--- program FrameL (robot ABB IRB 1300-10/1.15) ---
  Smooth(1)
  Set speed (1000.0 mm/s)
  Set Ref.: FrameL
  Set Tool: Generic Paint Sprayer
  Show Generic Paint Sprayer
  MoveJ 1 to (-13.41, 234.2, 55.45) mm, rotated rx -20.36 ry -7.23 rz -177.33 deg; joints [77.348, 64.389, -177.634, -26.013, 92.152, 94.605, 581.087, 3508.568, 217.224]
  MoveL 2 to (-13.41, 234.2, 55.45) mm, rotated rx -20.36 ry -7.23 rz -177.33 deg; joints [77.348, 64.389, -177.634, -26.013, 92.152, 94.605, 581.087, 3508.568, 217.224]
  MoveL 3 to (0, 200, 148.46) mm, rotated rx -20.36 ry -7.23 rz -177.33 deg; joints [77.348, 64.389, -177.634, -26.013, 92.152, 94.605, 594.495, 3417.935, 257.297]
  MoveL 4 to (0, 200, 148.46) mm, rotated rx -20.36 ry -7.23 rz -177.33 deg; joints [77.348, 64.389, -177.634, -26.013, 92.152, 94.605, 594.495, 3417.935, 257.297]
  Set speed (20.0 mm/s)
  MoveL 5 to (0, 100, 118.49) mm, rotated rx -13.25 ry -10.31 rz -177.59 deg; joints [77.348, 64.389, -177.469, -28.671, 97.668, 89.928, 571.606, 3460.539, 412.588]
  MoveL 6 to (0, 0, 100.67) mm, rotated rx -6.84 ry -13.03 rz -178.45 deg; joints [77.348, 64.389, -174.962, -31.186, 100.159, 86.521, 548.69, 3498.334, 553.088]
  Set speed (1000.0 mm/s)
  MoveL 7 to (0, 0, 100.67) mm, rotated rx -6.84 ry -13.03 rz -178.45 deg; joints [77.348, 64.389, -174.962, -31.186, 100.159, 86.521, 548.69, 3498.334, 553.088]
  MoveL 8 to (-22.71, 11.29, 3.94) mm, rotated rx -6.84 ry -13.03 rz -178.45 deg; joints [77.348, 64.389, -174.962, -31.186, 100.159, 86.521, 525.985, 3594.145, 535.636]
  Set speed (1000.0 mm/s)
  MoveL 9 to (70.65, -10.26, -4.8) mm, rotated rx 5.9 ry -2.48 rz 179.74 deg; joints [77.348, 64.389, -174.821, -21.333, 111.034, 81.501, 703.855, 3665.753, 651.653]
  MoveL 10 to (75, 0, 94.57) mm, rotated rx 5.9 ry -2.48 rz 179.74 deg; joints [77.348, 64.389, -174.821, -21.333, 111.034, 81.501, 708.205, 3565.924, 647.765]
  MoveL 11 to (75, 0, 94.57) mm, rotated rx 5.9 ry -2.48 rz 179.74 deg; joints [77.348, 64.389, -174.821, -21.333, 111.034, 81.501, 708.205, 3565.924, 647.765]
  Set speed (20.0 mm/s)
  MoveL 12 to (75, 100, 105.84) mm, rotated rx -14.61 ry -8.15 rz -177.88 deg; joints [77.348, 64.389, -193.763, -28.349, 111.034, 83.397, 684.859, 3386.076, 469.826]
  MoveL 13 to (75, 200, 138.19) mm, rotated rx -20.78 ry -6.55 rz -177.52 deg; joints [77.348, 76.516, -210, -27.07, 109.939, 85.836, 691.874, 3355.461, 460.291]
  Set speed (1000.0 mm/s)
  MoveL 14 to (75, 200, 138.19) mm, rotated rx -20.78 ry -6.55 rz -177.52 deg; joints [77.348, 76.516, -210, -27.07, 109.939, 85.836, 691.874, 3355.461, 460.291]
  MoveL 15 to (62.81, 234.98, 45.3) mm, rotated rx -20.78 ry -6.55 rz -177.52 deg; joints [77.348, 76.516, -210, -27.07, 109.939, 85.836, 679.685, 3445.924, 419.452]
  Set speed (1000.0 mm/s)
  MoveL 16 to (140.54, 234.66, 37.09) mm, rotated rx -20.96 ry 2.05 rz -159.4 deg; joints [79.127, 64.389, -196.024, -25.91, 117.994, 103.69, 801.481, 3466.335, 363.631]
  MoveL 17 to (150, 200, 130.42) mm, rotated rx -20.46 ry -5.09 rz -178.1 deg; joints [77.975, 76.516, -210, -26.014, 110.07, 85.836, 783.768, 3371.959, 458.597]
  MoveL 18 to (150, 200, 130.42) mm, rotated rx -20.46 ry -5.09 rz -178.1 deg; joints [77.975, 76.516, -210, -26.014, 110.07, 85.836, 783.768, 3371.959, 458.597]
  Set speed (20.0 mm/s)
  MoveL 19 to (150, 100, 95.81) mm, rotated rx -14.52 ry -5.16 rz -178.67 deg; joints [78.49, 76.516, -204.809, -26.013, 110.07, 84.398, 782.658, 3457.631, 573.254]
  MoveL 20 to (150, 0, 90.12) mm, rotated rx -1 ry -3.22 rz -179.94 deg; joints [78.49, 76.516, -192.395, -23.234, 110.07, 82.619, 785.471, 3572.863, 723.632]
  Set speed (1000.0 mm/s)
  MoveL 21 to (150, 0, 90.12) mm, rotated rx -1 ry -3.22 rz -179.94 deg; joints [78.49, 76.516, -192.395, -23.234, 110.07, 82.619, 785.471, 3572.863, 723.632]
  MoveL 22 to (144.37, 1.74, -9.71) mm, rotated rx -1 ry -3.22 rz -179.94 deg; joints [78.49, 76.516, -192.395, -23.234, 110.07, 82.619, 779.846, 3672.375, 715.52]
  Set speed (1000.0 mm/s)
  MoveL 23 to (196.55, 1, -12.04) mm, rotated rx -0.57 ry -1.97 rz -179.98 deg; joints [78.49, 76.516, -192.395, -21.96, 110.583, 82.834, 842.544, 3680.443, 719.238]
  MoveL 24 to (200, 0, 87.89) mm, rotated rx -0.57 ry -1.97 rz -179.98 deg; joints [78.49, 76.516, -192.395, -21.96, 110.583, 82.834, 845.989, 3580.776, 726.621]
  MoveL 25 to (200, 0, 87.89) mm, rotated rx -0.57 ry -1.97 rz -179.98 deg; joints [78.49, 76.516, -192.395, -21.96, 110.583, 82.834, 845.989, 3580.776, 726.621]
  Set speed (20.0 mm/s)
  MoveL 26 to (200, 100, 91.43) mm, rotated rx -14.97 ry -4.02 rz -178.93 deg; joints [78.49, 76.516, -205.685, -24.868, 110.583, 84.715, 843.258, 3461.359, 572.07]
  MoveL 27 to (200, 200, 126.09) mm, rotated rx -20.82 ry -4.07 rz -178.45 deg; joints [78.116, 76.516, -210, -24.986, 109.784, 86.361, 843.53, 3379.737, 453.356]
  Set speed (1000.0 mm/s)
  MoveL 28 to (200, 200, 126.09) mm, rotated rx -20.82 ry -4.07 rz -178.45 deg; joints [78.116, 76.516, -210, -24.986, 109.784, 86.361, 843.53, 3379.737, 453.356]
  MoveL 29 to (192.4, 235.34, 32.86) mm, rotated rx -20.82 ry -4.07 rz -178.45 deg; joints [78.116, 76.516, -210, -24.986, 109.784, 86.361, 835.932, 3470.525, 412.127]

--- program FrameR (robot ABB IRB 1300-10/1.15) ---
  Smooth(1)
  Set speed (1000.0 mm/s)
  Set Ref.: FrameR
  Set Tool: Generic Paint Sprayer
  Show Generic Paint Sprayer
  MoveJ 1 to (-1567.41, -947.44, 561.3) mm, rotated rx 116.18 ry 8.07 rz 164.06 deg; joints [-18.613, 70.643, -160.975, 159.818, -72.367, 68.936, 14.365, 240.215, 405.979]
  MoveL 2 to (-1567.41, -947.44, 561.3) mm, rotated rx 116.18 ry 8.07 rz 164.06 deg; joints [-18.613, 70.643, -160.975, 159.818, -72.367, 68.936, 14.365, 240.215, 405.979]
  MoveL 3 to (-1536.8, -862.85, 517.62) mm, rotated rx 116.18 ry 8.07 rz 164.06 deg; joints [-18.613, 70.643, -160.975, 159.818, -72.367, 68.936, 44.975, 324.8, 449.664]
  MoveL 4 to (-1536.8, -862.85, 517.62) mm, rotated rx 116.18 ry 8.07 rz 164.06 deg; joints [-18.613, 70.643, -160.975, 159.818, -72.367, 68.936, 44.975, 324.8, 449.664]
  Set speed (200.0 mm/s)
  MoveL 5 to (-1511.42, -864.68, 530.96) mm, rotated rx 117.6 ry 7.57 rz 165.86 deg; joints [-18.613, 70.643, -160.975, 158.345, -70.921, 68.501, 83.279, 316.894, 423.259]
  MoveL 6 to (-1485.52, -866.25, 542.73) mm, rotated rx 119.49 ry 6.77 rz 168.23 deg; joints [-18.613, 70.643, -160.989, 156.392, -68.942, 68.006, 127.136, 308.433, 393.799]
  MoveL 7 to (-1458.84, -867.56, 552.68) mm, rotated rx 120.63 ry 6.22 rz 169.63 deg; joints [-18.608, 70.645, -160.989, 155.208, -67.701, 67.76, 164.896, 303.689, 373.04]
  MoveL 8 to (-1431.63, -868.61, 560.79) mm, rotated rx 121.87 ry 5.07 rz 171.91 deg; joints [-18.608, 70.645, -161.394, 153.058, -66.382, 67.76, 214.467, 295.937, 351.142]
  MoveL 9 to (-1403.9, -869.65, 567.06) mm, rotated rx 122.48 ry 4.46 rz 173.04 deg; joints [-18.608, 70.645, -161.65, 151.982, -65.747, 67.76, 254.1, 292.049, 337.984]
  MoveL 10 to (-1375.91, -870.7, 571.77) mm, rotated rx 122.85 ry 3.63 rz 174.4 deg; joints [-18.607, 70.645, -162.511, 150.654, -65.699, 67.76, 300.795, 287.554, 327.831]
  MoveL 11 to (-1347.65, -871.48, 574.39) mm, rotated rx 123.43 ry 2.18 rz 176.71 deg; joints [-18.607, 70.645, -163.965, 148.372, -65.568, 67.76, 361.589, 281.477, 316.442]
  MoveL 12 to (-1319.14, -872.53, 575.44) mm, rotated rx 123.01 ry 1.1 rz 178.31 deg; joints [-18.607, 70.645, -164.386, 146.346, -65.568, 68.646, 409.222, 272.173, 314.488]
  MoveL 13 to (-1290.62, -873.32, 574.39) mm, rotated rx 122.75 ry 0.03 rz 179.95 deg; joints [-18.607, 70.645, -164.966, 144.398, -65.568, 69.295, 458.433, 264.711, 313.88]
  MoveL 14 to (-1262.63, -874.1, 571.51) mm, rotated rx 121.5 ry -0.87 rz -178.58 deg; joints [-18.607, 70.645, -164.966, 142.218, -65.996, 70.794, 501.334, 252.628, 322.32]
  MoveL 15 to (-1234.64, -874.62, 567.06) mm, rotated rx 119.59 ry -1.16 rz -177.95 deg; joints [-18.607, 70.645, -164.966, 140.919, -67.366, 72.2, 535.411, 241.481, 339.756]
  MoveL 16 to (-1207.43, -875.41, 561.05) mm, rotated rx 117.47 ry -1.89 rz -176.36 deg; joints [-18.607, 70.645, -164.966, 138.54, -68.641, 74.029, 577.946, 226.627, 358.999]
  MoveL 17 to (-1181.01, -875.67, 553.72) mm, rotated rx 114.97 ry -2.36 rz -174.95 deg; joints [-18.607, 70.645, -164.966, 136.4, -70.403, 75.823, 617.522, 212.418, 383.818]
  MoveL 18 to (-1155.11, -876.19, 544.57) mm, rotated rx 113.17 ry -2.69 rz -173.75 deg; joints [-18.607, 70.645, -164.966, 134.745, -71.68, 77.07, 654.392, 202.078, 405.856]
  MoveL 19 to (-1130.25, -876.46, 534.1) mm, rotated rx 110.41 ry -2.6 rz -173.06 deg; joints [-18.607, 70.645, -164.966, 133.557, -74.022, 78.489, 684.783, 190.934, 438.633]
  MoveL 20 to (-1106.18, -876.46, 522.33) mm, rotated rx 107.69 ry -2.35 rz -172.66 deg; joints [-18.607, 70.645, -164.966, 132.771, -76.442, 79.73, 711.467, 182.061, 473.425]
  MoveL 21 to (-1082.9, -876.72, 508.72) mm, rotated rx 105 ry -2.28 rz -171.55 deg; joints [-18.607, 70.645, -164.966, 131.287, -78.713, 81.041, 744.285, 172.206, 509.473]
  MoveL 22 to (-1060.66, -876.46, 493.81) mm, rotated rx 102.34 ry -1.62 rz -172.64 deg; joints [-18.368, 70.645, -164.966, 131.892, -81.381, 81.898, 754.662, 172.209, 549.165]
  MoveL 23 to (-1048.89, -876.46, 484.92) mm, rotated rx 101.61 ry -1.74 rz -171.59 deg; joints [-18.368, 70.645, -164.966, 130.744, -81.892, 82.332, 775.999, 168.058, 563.788]
  Set speed (1000.0 mm/s)
  MoveL 24 to (-1048.89, -876.46, 484.92) mm, rotated rx 101.61 ry -1.74 rz -171.59 deg; joints [-18.368, 70.645, -164.966, 130.744, -81.892, 82.332, 775.999, 168.058, 563.788]
  MoveL 25 to (-1033.96, -973.27, 505.03) mm, rotated rx 101.61 ry -1.74 rz -171.59 deg; joints [-18.368, 70.645, -164.966, 130.744, -81.892, 82.332, 790.935, 71.246, 543.68]
  Set speed (1000.0 mm/s)
  MoveL 26 to (-1620.34, -905.96, 635.31) mm, rotated rx 95.09 ry -1.66 rz -161.98 deg; joints [-23.506, 70.645, -168.71, 125.797, -89.471, 82.332, 337.544, 71.246, 474.728]
  MoveL 27 to (-1651.39, -811.31, 626.45) mm, rotated rx 95.09 ry -1.66 rz -161.98 deg; joints [-23.507, 70.645, -168.71, 125.798, -89.471, 82.332, 306.493, 165.888, 483.588]
  MoveL 28 to (-1651.39, -811.31, 626.45) mm, rotated rx 95.09 ry -1.66 rz -161.98 deg; joints [-23.507, 70.645, -168.71, 125.798, -89.471, 82.332, 306.493, 165.888, 483.588]
  Set speed (200.0 mm/s)
  MoveL 29 to (-1645.89, -808.17, 640.32) mm, rotated rx 113.53 ry -8.08 rz -162.12 deg; joints [-23.507, 72.673, -168.71, 127.007, -69.184, 79.927, 306.494, 206.634, 309.416]
  MoveL 30 to (-1651.65, -799.02, 663.34) mm, rotated rx 121.42 ry -9.52 rz -164.85 deg; joints [-23.507, 72.673, -168.71, 130.57, -61.954, 76.902, 284.437, 252.951, 222.205]
  MoveL 31 to (-1666.56, -784.63, 693.42) mm, rotated rx 124.61 ry -9.92 rz -165.99 deg; joints [-23.507, 73.957, -168.71, 131.64, -58.294, 76.527, 250.715, 279.424, 178.795]
  MoveL 32 to (-1677.55, -774.95, 712.52) mm, rotated rx 126.3 ry -10.62 rz -165.92 deg; joints [-23.574, 73.957, -168.71, 131.661, -56.497, 76.164, 244.342, 297.996, 145.936]
  MoveL 33 to (-1683.83, -769.72, 722.72) mm, rotated rx 125.13 ry -10.25 rz -165.82 deg; joints [-23.558, 73.957, -169.107, 131.661, -57.93, 76.164, 239.386, 297.902, 145.355]
  MoveL 34 to (-1683.83, -769.72, 722.72) mm, rotated rx 171.16 ry 2.79 rz 179.57 deg; joints [-36.296, 73.957, -189.291, 194.827, -57.93, 27.33, 239.385, 619.77, 42.153]
  MoveL 35 to (-1643.8, -776.52, 722.72) mm, rotated rx 171.27 ry 13.42 rz 177.96 deg; joints [-36.914, 73.957, -189.291, 200.842, -67.394, 24.825, 197.215, 619.774, 96.315]
  MoveL 36 to (-1607.96, -779.4, 730.31) mm, rotated rx 167.94 ry 10.28 rz 177.82 deg; joints [-33.158, 73.957, -189.291, 194.194, -66.22, 26.961, 238.044, 614.627, 76.195]
  MoveL 37 to (-1574.47, -782.8, 735.54) mm, rotated rx 162.76 ry 12.18 rz 176.26 deg; joints [-33.158, 73.957, -186.255, 192.105, -66.997, 30.46, 238.043, 566.815, 81.388]
  Set speed (1000.0 mm/s)
  MoveL 38 to (-1574.47, -782.8, 735.54) mm, rotated rx 162.76 ry 12.18 rz 176.26 deg; joints [-33.158, 73.957, -186.255, 192.105, -66.997, 30.46, 238.043, 566.815, 81.388]
  MoveL 39 to (-1596.51, -811.05, 828.9) mm, rotated rx 162.76 ry 12.18 rz 176.26 deg; joints [-33.158, 75.195, -187.492, 192.105, -66.997, 30.46, 213.238, 536.755, 0.003]
  Set speed (1000.0 mm/s)
  MoveL 40 to (-1593.63, -878.91, 757.51) mm, rotated rx 98.12 ry 1.45 rz 169.97 deg; joints [-33.158, 75.195, -183.445, 163.358, -101.211, 79.486, 213.238, 138.256, 406.615]
  MoveL 41 to (-1576.04, -781.49, 743.39) mm, rotated rx 98.12 ry 1.45 rz 169.97 deg; joints [-33.158, 75.195, -183.445, 163.358, -101.211, 79.486, 230.829, 235.678, 420.735]
  MoveL 42 to (-1576.04, -781.49, 743.39) mm, rotated rx 98.12 ry 1.45 rz 169.97 deg; joints [-33.158, 75.195, -183.445, 163.358, -101.211, 79.486, 230.829, 235.678, 420.735]
  Set speed (200.0 mm/s)
  MoveL 43 to (-1574.47, -782.27, 739.73) mm, rotated rx 97.18 ry 1.28 rz 169.93 deg; joints [-33.158, 75.195, -183.201, 163.264, -101.701, 80.152, 230.829, 233.1, 431.046]
  MoveL 44 to (-1571.6, -783.32, 735.54) mm, rotated rx 102.36 ry 2.06 rz 170.68 deg; joints [-33.158, 75.729, -183.201, 163.488, -97.124, 76.98, 234.295, 233.103, 398.064]
  MoveL 45 to (-1568.19, -785.41, 730.05) mm, rotated rx 108.49 ry 2.67 rz 172.07 deg; joints [-33.158, 76.713, -183.201, 163.595, -91.261, 73.401, 239.31, 233.102, 362.103]
  MoveL 46 to (-1563.75, -789.08, 722.2) mm, rotated rx 111.32 ry 2.84 rz 172.75 deg; joints [-33.158, 76.962, -183.201, 163.705, -88.725, 71.728, 246.486, 233.102, 349.55]
  MoveL 47 to (-1557.21, -794.31, 711.74) mm, rotated rx 113.21 ry 2.87 rz 173.35 deg; joints [-33.158, 76.962, -183.201, 163.673, -87.145, 70.589, 257.356, 231.07, 345.118]
  MoveL 48 to (-1543.86, -806.08, 689.5) mm, rotated rx 112.74 ry 3 rz 172.89 deg; joints [-32.822, 76.962, -182.72, 163.673, -87.145, 70.89, 262.386, 220.973, 370.252]
  MoveL 49 to (-1538.37, -810.27, 681.65) mm, rotated rx 112.52 ry 3.31 rz 172.07 deg; joints [-32.75, 76.961, -182.72, 164.391, -87.566, 70.949, 260.5, 220.973, 381.211]
  MoveL 50 to (-1531.83, -814.19, 674.59) mm, rotated rx 113.2 ry 2.69 rz 173.74 deg; joints [-32.75, 76.961, -182.72, 162.867, -86.528, 70.657, 281.259, 210.637, 380.287]
  MoveL 51 to (-1524.51, -817.85, 668.31) mm, rotated rx 113.92 ry 2.93 rz 173.42 deg; joints [-32.75, 76.961, -182.72, 163.435, -86.107, 70.178, 285.413, 211.149, 381.936]
  MoveL 52 to (-1516.4, -821.25, 663.08) mm, rotated rx 112.76 ry 3.01 rz 172.86 deg; joints [-32.542, 76.961, -182.257, 163.435, -86.681, 70.937, 285.42, 206.557, 395.395]
  MoveL 53 to (-1507.76, -824.39, 658.89) mm, rotated rx 109.21 ry 2.91 rz 171.71 deg; joints [-32.402, 76.916, -182.257, 163.435, -89.666, 73.068, 285.419, 199.674, 427.279]
  MoveL 54 to (-1498.61, -826.75, 656.01) mm, rotated rx 109.9 ry 2.54 rz 173.03 deg; joints [-32.402, 76.916, -182.258, 162.277, -88.785, 72.69, 305.443, 192.437, 423.021]
  MoveL 55 to (-1489.19, -828.84, 654.18) mm, rotated rx 107.78 ry 2.44 rz 172.43 deg; joints [-32.365, 76.916, -181.423, 162.277, -89.745, 74.227, 305.447, 184.607, 439.56]
  MoveL 56 to (-1479.51, -830.41, 653.66) mm, rotated rx 108.96 ry 2.29 rz 173.36 deg; joints [-32.365, 76.916, -181.423, 161.636, -88.611, 73.537, 322.581, 181.509, 429.869]
  MoveL 57 to (-1428.23, -836.69, 652.87) mm, rotated rx 112.95 ry 1.82 rz 175.71 deg; joints [-32.365, 76.916, -181.424, 160.346, -84.86, 71.308, 393.108, 176.138, 396.691]
  MoveL 58 to (-1385.33, -840.88, 652.09) mm, rotated rx 113.89 ry 1.35 rz 176.95 deg; joints [-32.365, 76.916, -181.424, 159.328, -83.722, 70.904, 447.029, 169.407, 388.191]
  MoveL 59 to (-1341.9, -844.02, 651.57) mm, rotated rx 113.18 ry 1.15 rz 177.32 deg; joints [-32.365, 76.916, -181.269, 158.734, -84.013, 71.415, 492.999, 161.611, 393.106]
  MoveL 60 to (-1314.69, -845.58, 651.04) mm, rotated rx 113.65 ry 1.17 rz 177.34 deg; joints [-32.249, 77.105, -181.269, 158.734, -83.449, 71.189, 518.198, 161.611, 391.36]
  MoveL 61 to (-1305.01, -845.58, 652.35) mm, rotated rx 113.89 ry 1.18 rz 177.34 deg; joints [-32.235, 77.284, -181.269, 158.773, -83.092, 71.116, 526.446, 161.611, 389.548]
  MoveL 62 to (-1296.12, -844.28, 656.27) mm, rotated rx 112.25 ry 0.44 rz 178.92 deg; joints [-32.235, 77.284, -181.226, 156.661, -83.843, 72.256, 549.803, 150.421, 395.544]
  MoveL 63 to (-1288.27, -842.18, 662.29) mm, rotated rx 109.89 ry -0.2 rz -179.46 deg; joints [-32.235, 77.284, -181.225, 154.389, -85.281, 73.661, 572.589, 138.737, 405.907]
  MoveL 64 to (-1282.25, -839.04, 669.88) mm, rotated rx 113.65 ry 0.48 rz 178.91 deg; joints [-32.235, 77.286, -181.23, 157.059, -82.712, 71.482, 563.484, 160.403, 371.001]
  MoveL 65 to (-1278.85, -835.12, 679.03) mm, rotated rx 113.65 ry 0.13 rz 179.7 deg; joints [-32.317, 77.286, -181.23, 156.309, -82.452, 71.61, 574.687, 160.404, 360.488]
  MoveL 66 to (-1277.54, -830.93, 688.71) mm, rotated rx 113.66 ry 0.65 rz 178.52 deg; joints [-32.317, 77.71, -181.23, 157.531, -82.452, 71.603, 561.67, 167.436, 355.878]
  MoveL 67 to (-1279.11, -826.49, 698.39) mm, rotated rx 113.19 ry 1.66 rz 176.12 deg; joints [-32.317, 77.959, -181.23, 159.893, -83.38, 71.634, 536.353, 179.707, 355.876]
  MoveL 68 to (-1282.51, -822.82, 706.5) mm, rotated rx 112.01 ry 1.43 rz 176.46 deg; joints [-32.317, 77.951, -181.23, 159.203, -84.202, 72.371, 536.352, 177.924, 356.114]
  MoveL 69 to (-1287.22, -818.9, 715.4) mm, rotated rx 109.18 ry 1.43 rz 175.91 deg; joints [-32.485, 77.234, -181.23, 159.196, -87.271, 73.747, 533.82, 177.924, 364.649]
  MoveL 70 to (-1291.67, -816.02, 722.99) mm, rotated rx 105.18 ry 1.04 rz 176.17 deg; joints [-32.485, 77.049, -181.23, 157.979, -90.559, 75.959, 533.82, 170.277, 387.037]
  MoveL 71 to (-1294.81, -814.45, 728.74) mm, rotated rx 100.47 ry 0.65 rz 176.47 deg; joints [-32.485, 77.049, -181.224, 156.739, -94.298, 78.535, 533.825, 161.41, 419.179]
  MoveL 72 to (-1297.16, -813.67, 732.67) mm, rotated rx 97.77 ry 0.62 rz 175.5 deg; joints [-32.485, 77.049, -181.224, 157.267, -96.675, 80.1, 523.529, 162.939, 438.079]
  MoveL 73 to (-1298.99, -813.14, 736.07) mm, rotated rx 89.91 ry -0.01 rz 175.41 deg; joints [-32.485, 76.771, -181.224, 156.398, -103.36, 84.313, 523.529, 160.679, 497.487]
  Set speed (1000.0 mm/s)
  MoveL 74 to (-1298.99, -813.14, 736.07) mm, rotated rx 89.91 ry -0.01 rz 175.41 deg; joints [-32.485, 76.771, -181.224, 156.398, -103.36, 84.313, 523.529, 160.679, 497.487]
  MoveL 75 to (-1306.99, -912.82, 735.92) mm, rotated rx 89.91 ry -0.01 rz 175.41 deg; joints [-32.485, 76.771, -181.224, 156.398, -103.36, 84.313, 515.53, 61, 497.634]
  Set speed (1000.0 mm/s)
  MoveL 76 to (-1277.26, -812.46, 899.51) mm, rotated rx 130.43 ry 1.94 rz 177.73 deg; joints [-32.485, 82.485, -181.224, 164.314, -65.405, 62.278, 515.529, 241.607, 65.66]
  MoveL 77 to (-1272.05, -736.49, 834.7) mm, rotated rx 130.43 ry 1.94 rz 177.73 deg; joints [-32.485, 82.485, -181.224, 164.314, -65.405, 62.278, 520.743, 317.58, 130.474]
  MoveL 78 to (-1272.05, -736.49, 834.7) mm, rotated rx 130.43 ry 1.94 rz 177.73 deg; joints [-32.485, 82.485, -181.224, 164.314, -65.405, 62.278, 520.743, 317.58, 130.474]
  Set speed (200.0 mm/s)
  MoveL 79 to (-1313.64, -732.57, 835.74) mm, rotated rx 131.13 ry 1.86 rz 177.87 deg; joints [-32.486, 82.485, -181.225, 164.465, -64.816, 61.836, 480.451, 324.806, 124.566]
  MoveL 80 to (-1348.7, -729.17, 836.53) mm, rotated rx 131.51 ry 2.46 rz 177.23 deg; joints [-32.486, 82.585, -181.206, 165.473, -64.817, 61.212, 437.294, 332.811, 124.566]
  MoveL 81 to (-1370.15, -726.81, 837.05) mm, rotated rx 131.03 ry 2.25 rz 177.41 deg; joints [-32.486, 82.375, -181.206, 165.02, -65.244, 61.624, 419.632, 332.534, 124.566]
  MoveL 82 to (-1401.81, -723.67, 837.57) mm, rotated rx 132.04 ry 2.5 rz 177.23 deg; joints [-32.486, 82.375, -181.206, 165.762, -64.645, 60.747, 385.483, 342.305, 118.589]
  MoveL 83 to (-1441.84, -719.23, 838.1) mm, rotated rx 133.18 ry 2.93 rz 176.89 deg; joints [-32.49, 82.375, -181.783, 166.881, -64.645, 59.499, 344.476, 357.293, 113.753]
  MoveL 84 to (-1485.26, -713.73, 838.88) mm, rotated rx 133.65 ry 3 rz 176.86 deg; joints [-32.492, 82.375, -182.089, 167.201, -64.645, 59.035, 302.34, 366.865, 110.952]
  MoveL 85 to (-1528.43, -707.71, 839.4) mm, rotated rx 134.21 ry 4.21 rz 175.68 deg; joints [-32.492, 82.375, -181.644, 169.049, -64.645, 57.959, 242.645, 380.514, 111.34]
  MoveL 86 to (-1562.18, -702.74, 839.67) mm, rotated rx 135.2 ry 4.73 rz 175.31 deg; joints [-32.493, 82.375, -181.868, 170.148, -64.51, 56.845, 205.151, 394.369, 107.799]
  MoveL 87 to (-1610.05, -694.63, 839.67) mm, rotated rx 135.22 ry 5.08 rz 174.98 deg; joints [-32.493, 82.375, -181.638, 170.602, -64.511, 56.652, 152, 403.576, 108.755]
  MoveL 88 to (-1652.17, -686.26, 839.67) mm, rotated rx 135.73 ry 5.47 rz 174.69 deg; joints [-32.493, 82.375, -181.727, 171.316, -64.511, 56.005, 106.555, 417.077, 107.647]
  MoveL 89 to (-1691.68, -677.63, 839.67) mm, rotated rx 136.03 ry 5.85 rz 174.38 deg; joints [-32.493, 82.383, -181.727, 171.926, -64.56, 55.539, 63.117, 429.319, 107.647]
  MoveL 90 to (-1724.9, -670.56, 838.1) mm, rotated rx 136.82 ry 6.43 rz 174 deg; joints [-32.493, 82.383, -181.876, 172.973, -64.56, 54.549, 25.38, 444.226, 107.518]
  MoveL 91 to (-1758.39, -661.41, 836.26) mm, rotated rx 135.23 ry 8 rz 172.14 deg; joints [-34.724, 80.46, -181.876, 176.549, -68.763, 55.099, 0.002, 444.226, 110.987]
  Set speed (1000.0 mm/s)
  MoveL 92 to (-1758.39, -661.41, 836.26) mm, rotated rx 135.23 ry 8 rz 172.14 deg; joints [-34.724, 80.46, -181.876, 176.549, -68.763, 55.099, 0.002, 444.226, 110.987]
  MoveL 93 to (-1777.81, -729.83, 906.56) mm, rotated rx 135.23 ry 8 rz 172.14 deg; joints [-34.724, 80.46, -185.22, 176.62, -72.101, 54.888, 0, 389.269, 48.578]
  Set speed (1000.0 mm/s)
  MoveL 94 to (892.89, -973.97, 160.56) mm, rotated rx 74.09 ry -79.65 rz -165.04 deg; joints [-50.625, 101.986, -183.176, 143.958, -56.047, 174.635, 2943.702, -296.83, 1100]
  MoveL 95 to (894.12, -874.1, 165.49) mm, rotated rx 74.09 ry -79.65 rz -165.04 deg; joints [-50.625, 102.249, -183.176, 143.853, -55.834, 174.822, 2944.041, -198.044, 1097.78]
  MoveL 96 to (894.12, -874.1, 165.49) mm, rotated rx 74.09 ry -79.65 rz -165.04 deg; joints [-50.625, 102.249, -183.176, 143.853, -55.834, 174.822, 2944.041, -198.044, 1097.78]
  Set speed (200.0 mm/s)
  MoveL 97 to (897.25, -874.89, 176.21) mm, rotated rx 65.87 ry -79.15 rz -157.31 deg; joints [-50.572, 102.13, -183.176, 144.306, -57.481, 174.822, 2944.041, -202.933, 1099.813]
  MoveL 98 to (899.87, -876.46, 192.17) mm, rotated rx 61.84 ry -78.73 rz -152.65 deg; joints [-50.572, 102.13, -183.176, 143.646, -58.425, 174.912, 2952.705, -207.84, 1091.736]
  MoveL 99 to (903.01, -878.29, 209.44) mm, rotated rx 62.04 ry -78.65 rz -151.92 deg; joints [-50.572, 102.13, -183.176, 142.694, -58.517, 174.948, 2963.908, -210.297, 1074.532]
  MoveL 100 to (906.93, -880.12, 229.58) mm, rotated rx 62.24 ry -78.57 rz -151.18 deg; joints [-50.572, 102.13, -183.176, 141.745, -58.61, 174.982, 2975.895, -212.626, 1054.448]
  MoveL 101 to (912.69, -881.95, 251.82) mm, rotated rx 63.48 ry -78.61 rz -151.46 deg; joints [-50.572, 102.13, -183.22, 140.789, -58.506, 174.982, 2989.943, -213.842, 1030.144]
  MoveL 102 to (920.28, -883.78, 275.36) mm, rotated rx 64.54 ry -78.72 rz -152.5 deg; joints [-50.571, 102.13, -183.221, 140.765, -58.272, 174.982, 2997.54, -214.928, 1004.496]
  MoveL 103 to (929.69, -885.35, 299.69) mm, rotated rx 65.62 ry -78.83 rz -153.56 deg; joints [-50.545, 102.13, -183.227, 140.714, -58.045, 174.982, 3006.729, -215.496, 978.065]
  MoveL 104 to (940.68, -886.66, 324.29) mm, rotated rx 66.79 ry -78.9 rz -154.23 deg; joints [-50.519, 102.13, -183.265, 140.199, -57.891, 174.982, 3021.693, -215.76, 951.388]
  MoveL 105 to (953.5, -887.97, 348.36) mm, rotated rx 85.13 ry -19.62 rz -174.48 deg; joints [0, 44.016, -168.118, 113.546, -98.533, 78.32, 3060.514, 351.718, 637.921]
  MoveL 106 to (968.15, -889.01, 371.64) mm, rotated rx 85.13 ry -19.62 rz -174.48 deg; joints [0, 44.016, -168.118, 113.546, -98.533, 78.32, 3075.164, 350.671, 614.638]
  MoveL 107 to (984.11, -889.8, 393.88) mm, rotated rx 84.63 ry -19.58 rz -174.31 deg; joints [0, 44.835, -168.118, 113.424, -98.568, 79.239, 3080.491, 349.61, 598.511]
  MoveL 108 to (1001.38, -890.32, 415.07) mm, rotated rx 85.13 ry -19.62 rz -174.48 deg; joints [0.001, 44.853, -168.118, 113.658, -98.197, 79.096, 3097.541, 349.369, 573.162]
  MoveL 109 to (1020.21, -890.58, 435.21) mm, rotated rx 84.63 ry -19.58 rz -174.31 deg; joints [0.001, 45.265, -168.118, 113.481, -98.396, 79.637, 3111.032, 348.831, 558.239]
  MoveL 110 to (1040.1, -890.84, 453.79) mm, rotated rx 84.38 ry -19.55 rz -174.23 deg; joints [0.001, 45.523, -168.118, 113.402, -98.476, 79.957, 3127.571, 348.445, 542.424]
  MoveL 111 to (1066.78, -890.84, 475.24) mm, rotated rx 84.63 ry -19.58 rz -174.31 deg; joints [0.001, 45.532, -168.118, 113.517, -98.289, 79.885, 3154.15, 348.57, 518.893]
  MoveL 112 to (1095.03, -890.58, 494.6) mm, rotated rx 85.13 ry -19.62 rz -174.48 deg; joints [0.001, 45.549, -168.118, 113.748, -97.917, 79.739, 3182.208, 349.108, 495.375]
  MoveL 113 to (1124.86, -890.06, 511.6) mm, rotated rx 85.38 ry -19.72 rz -175.5 deg; joints [0.001, 45.558, -168.118, 114.693, -98.158, 79.939, 3203.662, 352.782, 476.029]
  MoveL 114 to (1155.99, -889.54, 525.99) mm, rotated rx 85.88 ry -19.72 rz -175.19 deg; joints [0, 45.573, -168.118, 114.51, -97.577, 79.649, 3238.754, 352.115, 457.625]
  MoveL 115 to (1181.63, -888.75, 535.67) mm, rotated rx 86.12 ry -19.77 rz -175.75 deg; joints [0, 45.582, -168.118, 115.04, -97.607, 79.708, 3260.15, 354.598, 445.767]
  MoveL 116 to (1207.79, -887.97, 543.52) mm, rotated rx 86.62 ry -19.83 rz -176.38 deg; joints [0, 45.6, -168.118, 115.686, -97.454, 79.686, 3281.974, 357.321, 433.7]
  MoveL 117 to (1234.47, -887.18, 549.8) mm, rotated rx 86.87 ry -19.87 rz -176.94 deg; joints [0, 45.613, -168.118, 116.215, -97.485, 79.743, 3304.394, 359.899, 425.291]
  MoveL 118 to (1261.68, -886.4, 554.25) mm, rotated rx 87.62 ry -19.89 rz -176.72 deg; joints [0, 45.625, -168.118, 116.15, -96.728, 79.358, 3335.564, 359.768, 414.744]
  MoveL 119 to (1288.89, -885.35, 556.86) mm, rotated rx 88.12 ry -19.93 rz -177.36 deg; joints [0, 45.643, -168.118, 116.795, -96.582, 79.323, 3358.44, 362.895, 407.98]
  MoveL 120 to (1316.36, -884.57, 557.91) mm, rotated rx 88.12 ry -19.96 rz -178.3 deg; joints [0.004, 45.662, -168.118, 117.618, -97.006, 79.598, 3377.48, 366.981, 406.875]
  MoveL 121 to (1343.57, -883.78, 556.86) mm, rotated rx 88.12 ry -19.96 rz -178.3 deg; joints [0.004, 45.662, -168.118, 117.618, -97.006, 79.598, 3404.688, 367.766, 407.922]
  MoveL 122 to (1371.04, -883, 554.25) mm, rotated rx 87.87 ry -19.95 rz -178.21 deg; joints [-0.098, 45.662, -168.118, 117.592, -97.231, 79.716, 3432.156, 367.766, 412.586]
  MoveL 123 to (1398.24, -882.21, 549.8) mm, rotated rx 88.12 ry -19.96 rz -178.3 deg; joints [-0.098, 45.668, -168.118, 117.708, -97.052, 79.628, 3459.294, 368.802, 415]
  MoveL 124 to (1425.45, -881.43, 543.52) mm, rotated rx 88.87 ry -19.98 rz -178.56 deg; joints [-0.098, 45.682, -168.118, 118.055, -96.518, 79.362, 3486.317, 370.389, 415.176]
  MoveL 125 to (1452.4, -880.64, 535.67) mm, rotated rx 88.87 ry -19.98 rz -178.56 deg; joints [-0.098, 45.682, -168.118, 118.055, -96.518, 79.362, 3513.264, 371.174, 423.025]
  Set speed (1000.0 mm/s)
  MoveL 126 to (1452.4, -880.64, 535.67) mm, rotated rx 88.87 ry -19.98 rz -178.56 deg; joints [-0.098, 45.682, -168.118, 118.055, -96.518, 79.362, 3513.264, 371.174, 423.025]
  MoveL 127 to (1454.25, -980.61, 533.82) mm, rotated rx 88.87 ry -19.98 rz -178.56 deg; joints [-0.098, 45.682, -168.118, 118.055, -96.518, 79.362, 3515.111, 271.208, 424.873]
  Set speed (1000.0 mm/s)
  MoveL 128 to (1533.99, -926.46, 631.09) mm, rotated rx 138.74 ry -6.11 rz -174.67 deg; joints [-9.541, 61.146, -158.442, 135.819, -50.553, 59.636, 3391.215, 390.14, 48.578]
  MoveL 129 to (1519.9, -861.54, 556.34) mm, rotated rx 138.74 ry -6.11 rz -174.67 deg; joints [-9.541, 61.146, -158.442, 135.819, -50.553, 59.636, 3377.12, 455.057, 123.326]
  MoveL 130 to (1519.9, -861.54, 556.34) mm, rotated rx 138.74 ry -6.11 rz -174.67 deg; joints [-9.541, 61.146, -158.442, 135.819, -50.553, 59.636, 3377.12, 455.057, 123.326]
  Set speed (200.0 mm/s)
  MoveL 131 to (1489.29, -872.53, 551.89) mm, rotated rx 138.33 ry -11.97 rz -169.54 deg; joints [-9.406, 61.146, -158.442, 126.772, -46.624, 65.411, 3417.685, 437.6, 113.159]
  MoveL 132 to (1461.56, -873.05, 561.57) mm, rotated rx 139.84 ry -10.86 rz -170.96 deg; joints [-9.406, 61.146, -158.442, 129.677, -46.276, 63.079, 3373.678, 447.966, 98.005]
  MoveL 133 to (1433.04, -873.58, 569.68) mm, rotated rx 141.66 ry -9.37 rz -172.66 deg; joints [-9.406, 61.146, -158.442, 133.371, -46.012, 60.06, 3324.622, 461.468, 84.178]
  MoveL 134 to (1404.52, -874.36, 576.22) mm, rotated rx 143.33 ry -7.53 rz -174.43 deg; joints [-9.406, 61.146, -158.442, 137.332, -46.181, 56.838, 3272.974, 474.662, 74.367]
  MoveL 135 to (1375.22, -875.15, 580.67) mm, rotated rx 143.54 ry -5.51 rz -175.94 deg; joints [-9.406, 61.073, -158.442, 140.257, -47.619, 54.789, 3221.713, 478.344, 74.674]
  MoveL 136 to (1345.92, -875.93, 583.81) mm, rotated rx 143.06 ry -3.49 rz -177.38 deg; joints [-9.406, 61.217, -158.628, 142.541, -49.547, 53.504, 3169.819, 477.803, 82.221]
  MoveL 137 to (1316.1, -876.98, 585.12) mm, rotated rx 142.32 ry -2.18 rz -178.32 deg; joints [-9.406, 61.43, -158.905, 143.697, -51.125, 53.088, 3125.253, 474.44, 91.484]
  MoveL 138 to (1286.01, -877.76, 585.38) mm, rotated rx 140.67 ry -0.69 rz -179.43 deg; joints [-9.406, 61.887, -159.499, 144.523, -53.535, 53.312, 3077.773, 466.28, 109.947]
  MoveL 139 to (1255.14, -878.55, 584.07) mm, rotated rx 137.84 ry 0.78 rz 179.29 deg; joints [-9.406, 62.612, -160.443, 144.766, -56.841, 54.489, 3028.427, 451.799, 139.793]
  MoveL 140 to (1223.49, -879.07, 581.45) mm, rotated rx 134.73 ry 1.74 rz 178.25 deg; joints [-9.406, 63.328, -161.381, 144.461, -59.978, 56.161, 2983.148, 436.266, 171.527]
  MoveL 141 to (1190.26, -879.59, 578.05) mm, rotated rx 133.24 ry 1.97 rz 177.91 deg; joints [-9.406, 63.653, -161.807, 144.091, -61.33, 57.095, 2945.816, 428.197, 188.24]
  MoveL 142 to (1155.47, -879.59, 573.87) mm, rotated rx 131.24 ry 2.37 rz 177.3 deg; joints [-9.406, 64.059, -162.341, 143.811, -63.215, 58.243, 2904.186, 419.258, 210.694]
  MoveL 143 to (1117.01, -879.07, 569.16) mm, rotated rx 126.69 ry 2.59 rz 176.53 deg; joints [-9.406, 64.918, -163.475, 142.508, -67.052, 61.172, 2857.854, 398.451, 254.993]
  MoveL 144 to (1084.05, -880.38, 560) mm, rotated rx 121.8 ry 2.47 rz 176.03 deg; joints [-9.406, 65.478, -164.218, 140.911, -70.931, 64.405, 2821.001, 375.562, 303.776]
  MoveL 145 to (1052.39, -880.9, 553.98) mm, rotated rx 120.88 ry 0.65 rz 178.91 deg; joints [-9.834, 65.478, -164.218, 137.662, -70.306, 66.212, 2818.641, 353.715, 309.094]
  MoveL 146 to (1009.23, -879.33, 553.98) mm, rotated rx 119.04 ry 0.4 rz 179.27 deg; joints [-10.314, 65.479, -164.219, 137.039, -71.636, 67.57, 2780.014, 341.197, 321.813]
  Set speed (1000.0 mm/s)
  MoveL 147 to (1009.23, -879.33, 553.98) mm, rotated rx 119.04 ry 0.4 rz 179.27 deg; joints [-10.314, 65.479, -164.219, 137.039, -71.636, 67.57, 2780.014, 341.197, 321.813]
  MoveL 148 to (1007.78, -966.75, 602.53) mm, rotated rx 119.04 ry 0.4 rz 179.27 deg; joints [-10.314, 65.479, -164.219, 137.039, -71.636, 67.57, 2778.565, 253.784, 273.265]
  Set speed (1000.0 mm/s)
  MoveL 149 to (873.5, -880.28, 780.09) mm, rotated rx 138.11 ry -2.37 rz -177.88 deg; joints [-10.314, 69.754, -169.974, 142.569, -56.185, 54.961, 2673.473, 430.431, 0]
  MoveL 150 to (867.95, -813.67, 705.72) mm, rotated rx 138.11 ry -2.37 rz -177.88 deg; joints [-10.314, 69.754, -169.974, 142.569, -56.185, 54.961, 2667.932, 497.048, 74.374]
  MoveL 151 to (867.95, -813.67, 705.72) mm, rotated rx 138.11 ry -2.37 rz -177.88 deg; joints [-10.314, 69.754, -169.974, 142.569, -56.185, 54.961, 2667.932, 497.048, 74.374]
  Set speed (200.0 mm/s)
  MoveL 152 to (904.84, -813.67, 702.84) mm, rotated rx 138.4 ry -2.86 rz -177.46 deg; joints [-10.348, 69.754, -169.974, 142.156, -55.592, 55.078, 2710.558, 497.291, 73.781]
  MoveL 153 to (941.47, -813.41, 700.23) mm, rotated rx 139.78 ry -3.56 rz -176.99 deg; joints [-10.348, 69.694, -169.893, 142.201, -54.052, 54.45, 2754.696, 505.196, 65.514]
  MoveL 154 to (978.09, -813.14, 697.35) mm, rotated rx 140.31 ry -3.04 rz -177.48 deg; joints [-10.213, 69.694, -169.893, 143.129, -54.093, 53.594, 2784.707, 511.736, 67.35]
  MoveL 155 to (1014.72, -812.62, 694.47) mm, rotated rx 138.88 ry -3.15 rz -177.25 deg; joints [-10.213, 69.694, -169.893, 141.972, -54.989, 54.887, 2823.471, 502.14, 77.761]
  MoveL 156 to (1051.87, -812.1, 691.59) mm, rotated rx 137.92 ry -3.25 rz -177.07 deg; joints [-10.214, 69.694, -169.893, 141.188, -55.584, 55.745, 2862.315, 495.937, 85.751]
  MoveL 157 to (1090.33, -811.58, 688.45) mm, rotated rx 140.78 ry -3.42 rz -177.21 deg; joints [-10.214, 69.645, -169.825, 142.984, -53.446, 53.474, 2901.1, 515.702, 71.782]
  MoveL 158 to (1131.14, -810.79, 684.79) mm, rotated rx 141.73 ry -3.41 rz -177.31 deg; joints [-10.214, 69.629, -169.804, 143.689, -52.802, 52.645, 2941.325, 523.172, 70.224]
  MoveL 159 to (1175.09, -810.01, 680.6) mm, rotated rx 141.49 ry -3.86 rz -176.93 deg; joints [-10.214, 69.629, -169.804, 142.952, -52.605, 53.185, 2990.491, 521.26, 74.11]
  MoveL 160 to (1220.35, -808.96, 676.16) mm, rotated rx 141.93 ry -4.58 rz -176.42 deg; joints [-10.239, 69.647, -169.804, 142.399, -51.718, 53.352, 3043.49, 523.666, 73.879]
  MoveL 161 to (1265.35, -807.91, 671.45) mm, rotated rx 142.71 ry -3.96 rz -176.99 deg; joints [-10.076, 69.647, -169.803, 143.629, -51.673, 52.164, 3080.695, 533.169, 76.64]
  MoveL 162 to (1308.25, -806.6, 666.74) mm, rotated rx 142.43 ry -3.78 rz -177.1 deg; joints [-10.029, 69.733, -169.803, 143.556, -51.931, 52.336, 3120.743, 533.169, 84.07]
  MoveL 163 to (1347.49, -805.3, 662.29) mm, rotated rx 142.24 ry -4.83 rz -176.27 deg; joints [-10.206, 69.7, -169.758, 142.247, -51.221, 53.337, 3172.343, 529.258, 85.549]
  MoveL 164 to (1385.43, -803.73, 657.84) mm, rotated rx 141.75 ry -6.36 rz -175.01 deg; joints [-10.206, 69.7, -169.758, 139.926, -50.344, 54.95, 3228.058, 524.713, 87.591]
  MoveL 165 to (1429.12, -801.37, 651.83) mm, rotated rx 140.48 ry -6.48 rz -174.69 deg; joints [-10.206, 69.7, -169.758, 138.77, -51.128, 56.142, 3274.416, 517.767, 100.02]
  MoveL 166 to (1480.65, -797.97, 643.98) mm, rotated rx 140.88 ry -6.94 rz -174.39 deg; joints [-10.551, 69.337, -169.263, 138.71, -50.428, 56.337, 3331.85, 520.017, 100.585]
  MoveL 167 to (1525.91, -794.57, 636.39) mm, rotated rx 143.15 ry -7.95 rz -174.08 deg; joints [-10.551, 69.344, -169.263, 139.263, -48.057, 55.155, 3386.01, 538.846, 93.227]
  MoveL 168 to (1570.39, -790.38, 628.28) mm, rotated rx 142.96 ry -9.33 rz -173.02 deg; joints [-10.712, 69.33, -169.245, 137.427, -47.121, 56.529, 3446.772, 538.846, 98.189]
  MoveL 169 to (1604.14, -786.72, 621.48) mm, rotated rx 141.05 ry -10.48 rz -171.64 deg; joints [-10.712, 69.329, -169.243, 134.243, -47.573, 59.2, 3496.639, 527.838, 111.781]
  MoveL 170 to (1635.01, -782.8, 614.94) mm, rotated rx 141.92 ry -11.12 rz -171.41 deg; joints [-10.712, 69.3, -169.204, 134.121, -46.464, 59.025, 3533.455, 537.973, 111.775]
  MoveL 171 to (1664.04, -778.61, 608.4) mm, rotated rx 141.82 ry -12.17 rz -170.59 deg; joints [-11.054, 69.025, -168.829, 132.808, -45.717, 60.235, 3575.747, 537.973, 113.449]
  MoveL 172 to (1691.25, -774.16, 601.34) mm, rotated rx 142.72 ry -13.83 rz -169.68 deg; joints [-11.054, 69.024, -168.829, 131.288, -43.831, 61.04, 3620.345, 549.538, 112.01]
  MoveL 173 to (1717.15, -769.46, 594.01) mm, rotated rx 144.18 ry -14.24 rz -169.93 deg; joints [-11.054, 69.024, -168.829, 132.075, -42.496, 60.144, 3647.995, 565.322, 111.216]
  MoveL 174 to (1741.48, -764.22, 585.9) mm, rotated rx 143.22 ry -16.98 rz -167.69 deg; joints [-11.113, 69.024, -168.829, 127.258, -41.194, 63.853, 3705.229, 565.239, 118.706]
  MoveL 175 to (1763.46, -759.25, 577.79) mm, rotated rx 147.1 ry -20.86 rz -167.03 deg; joints [-11.113, 69.024, -168.829, 125.179, -35.697, 64.914, 3760.726, 604.805, 103.148]
  MoveL 176 to (1782.03, -754.81, 570.47) mm, rotated rx 149.6 ry -22.53 rz -167.33 deg; joints [-11.113, 69.024, -168.828, 125.124, -32.775, 64.732, 3791.331, 631.104, 98.349]
  MoveL 177 to (1797.47, -750.88, 563.66) mm, rotated rx 149.1 ry -22.89 rz -166.9 deg; joints [-11.207, 68.767, -168.479, 123.926, -32.856, 65.888, 3812.138, 631.104, 104.311]
  MoveL 178 to (1809.5, -747.74, 557.91) mm, rotated rx 149.34 ry -27.13 rz -164.88 deg; joints [-11.369, 68.485, -168.097, 116.582, -30.027, 72.314, 3867.977, 644.455, 104.311]
  MoveL 179 to (1819.44, -745.39, 552.94) mm, rotated rx 152.47 ry -25.62 rz -167.3 deg; joints [-11.369, 69.123, -168.963, 123.151, -28.77, 66.476, 3854.856, 665.831, 104.31]
  MoveL 180 to (1827.81, -743.03, 548.23) mm, rotated rx 155.32 ry -27.01 rz -168.21 deg; joints [-11.369, 69.123, -168.963, 123.836, -25.853, 65.81, 3871.651, 692.676, 99.167]
  Set speed (1000.0 mm/s)
  MoveL 181 to (1827.81, -743.03, 548.23) mm, rotated rx 155.32 ry -27.01 rz -168.21 deg; joints [-11.369, 69.123, -168.963, 123.836, -25.853, 65.81, 3871.651, 692.676, 99.167]
  MoveL 182 to (1876.74, -775.47, 629.18) mm, rotated rx 155.32 ry -27.01 rz -168.21 deg; joints [-11.369, 69.123, -168.963, 123.836, -25.853, 65.81, 3920.576, 660.235, 18.211]
  Set speed (1000.0 mm/s)
  MoveL 183 to (883.17, -844.02, 851.21) mm, rotated rx 124.16 ry -6.87 rz -170 deg; joints [-11.369, 72, -172.918, 127.917, -63.476, 67.716, 2763.544, 357.619, 25.596]
  MoveL 184 to (862.2, -763.7, 795.45) mm, rotated rx 124.16 ry -6.87 rz -170 deg; joints [-11.369, 71.999, -172.918, 127.917, -63.476, 67.715, 2742.569, 437.942, 81.346]
  MoveL 185 to (862.2, -763.7, 795.45) mm, rotated rx 124.16 ry -6.87 rz -170 deg; joints [-11.369, 71.999, -172.918, 127.917, -63.476, 67.715, 2742.569, 437.942, 81.346]
  Set speed (200.0 mm/s)
  MoveL 186 to (834.21, -757.94, 813.24) mm, rotated rx 125.41 ry -7.49 rz -169.6 deg; joints [-11.997, 71.344, -172.918, 128.596, -62.551, 66.897, 2728.773, 444.882, 47.939]
  MoveL 187 to (805.69, -752.19, 831.29) mm, rotated rx 128.43 ry -8.31 rz -169.68 deg; joints [-12.476, 70.429, -172.918, 130.342, -60.33, 64.815, 2714.571, 464.902, 0.024]
  MoveL 188 to (775.87, -745.91, 849.87) mm, rotated rx 128.95 ry -7.87 rz -170.38 deg; joints [-12.476, 72.403, -175.69, 131.734, -60.838, 63.479, 2676.515, 474.819, 0]
  MoveL 189 to (743.95, -739.37, 869.23) mm, rotated rx 130.21 ry -8.72 rz -169.84 deg; joints [-12.476, 75.224, -179.751, 131.973, -60.065, 62.154, 2654.218, 488.345, 0]
  MoveL 190 to (709.42, -732.04, 889.63) mm, rotated rx 133.19 ry -9.83 rz -169.7 deg; joints [-12.476, 79.053, -185.502, 133.645, -58.375, 59.225, 2632.238, 514.975, 0]
  MoveL 191 to (673.05, -724.2, 910.56) mm, rotated rx 134.82 ry -10.39 rz -169.71 deg; joints [-12.476, 81.857, -189.951, 134.999, -57.948, 57.058, 2605.927, 534.847, 0]
  MoveL 192 to (634.86, -716.35, 931.75) mm, rotated rx 135.84 ry -10.15 rz -170.29 deg; joints [-12.476, 84.07, -193.661, 136.805, -58.584, 54.965, 2569.677, 551.383, 0]
  MoveL 193 to (590.38, -706.67, 956.08) mm, rotated rx 134.93 ry -9.14 rz -170.95 deg; joints [-13.013, 85.36, -195.933, 138.055, -60.928, 54.432, 2520.708, 551.818, 0]
  MoveL 194 to (534.66, -694.63, 985.12) mm, rotated rx 133.18 ry -7.68 rz -171.9 deg; joints [-13.013, 86.447, -197.926, 138.708, -64.085, 54.194, 2454.494, 554.996, 0.002]
  MoveL 195 to (471.61, -681.29, 1016.78) mm, rotated rx 130.54 ry -5.99 rz -173.05 deg; joints [-13.013, 87.161, -199.282, 138.966, -67.883, 54.662, 2377.062, 555.261, 0.001]
  MoveL 196 to (405.16, -667.16, 1047.91) mm, rotated rx 124.82 ry -2.46 rz -176.48 deg; joints [-12.982, 84.421, -199.282, 140.33, -77.278, 54.915, 2286.095, 552.193, 2.626]
  MoveL 197 to (341.85, -654.08, 1076.43) mm, rotated rx 122.99 ry -1.83 rz -177.19 deg; joints [-12.982, 85.194, -200.802, 140.238, -79.759, 55.286, 2218.458, 559.632, 0.082]
  MoveL 198 to (288.22, -643.1, 1099.97) mm, rotated rx 124.74 ry -1.97 rz -177.17 deg; joints [-12.982, 87.676, -206.184, 141.414, -80.688, 52.498, 2181.903, 582.709, 0]
  MoveL 199 to (239.56, -634.46, 1118.81) mm, rotated rx 128.95 ry 13.04 rz -164.09 deg; joints [-31.64, 82.162, -208.59, 150.889, -96.953, 37.959, 2259.037, 439.327, 0]
  MoveL 200 to (190.9, -627.66, 1133.72) mm, rotated rx 126.76 ry 14.31 rz -165.51 deg; joints [-31.64, 82.162, -208.589, 150.719, -99.462, 38.725, 2200.517, 438.925, 6.01]
  MoveL 201 to (142.76, -622.17, 1145.75) mm, rotated rx 124.74 ry 15.48 rz -167.01 deg; joints [-31.64, 82.162, -208.589, 150.763, -101.829, 39.458, 2141.901, 439.363, 13.545]
  MoveL 202 to (95.15, -617.72, 1156.22) mm, rotated rx 136.3 ry 27.91 rz -149.96 deg; joints [-44.422, 91.876, -166.166, 151.842, -57.295, 47.859, 1940.01, 93.218, 0.016]
  MoveL 203 to (45.18, -613.53, 1165.11) mm, rotated rx 140.79 ry 25.55 rz -147.99 deg; joints [-44.422, 95.911, -166.166, 150.356, -49.393, 48.719, 1870.377, 97.394, 0.001]
  MoveL 204 to (-9.5, -609.09, 1172.7) mm, rotated rx 137.9 ry 28.6 rz -150.73 deg; joints [-44.443, 95.606, -166.166, 152.95, -53.361, 47.699, 1800.439, 91.784, 22.931]
  MoveL 205 to (-66.79, -605.42, 1178.72) mm, rotated rx 136.64 ry 29.48 rz -151.63 deg; joints [-44.443, 95.632, -166.201, 153.428, -54.7, 47.81, 1739.995, 91.323, 29.345]
  MoveL 206 to (-124.09, -602.02, 1183.43) mm, rotated rx 133.51 ry 31.81 rz -154.34 deg; joints [-44.443, 95.508, -166.201, 155.176, -58.15, 47.675, 1671.169, 87.512, 54.709]
  MoveL 207 to (-178.76, -599.41, 1187.09) mm, rotated rx 133.6 ry 31.93 rz -154.49 deg; joints [-44.443, 95.508, -166.201, 155.436, -58.161, 47.456, 1614.474, 90.776, 51.361]
  MoveL 208 to (-228.21, -597.31, 1189.97) mm, rotated rx 133.46 ry 31.71 rz -154.21 deg; joints [-44.589, 95.508, -166.201, 155.135, -58.103, 47.789, 1570.121, 90.265, 47.767]
  MoveL 209 to (-273.47, -595.74, 1192.06) mm, rotated rx 136.82 ry 29.2 rz -151.33 deg; joints [-44.658, 95.507, -166.2, 153.394, -54.499, 47.837, 1538.388, 99.677, 11.784]
  MoveL 210 to (-315.85, -594.17, 1193.89) mm, rotated rx 141.11 ry 27.24 rz -149.49 deg; joints [-44.658, 97.542, -166.2, 152.858, -48.762, 47.23, 1485.019, 109.494, 0]
  MoveL 211 to (-357.71, -592.87, 1194.94) mm, rotated rx 138.48 ry 28.97 rz -151.11 deg; joints [-44.658, 97.414, -166.2, 153.623, -51.59, 47.611, 1439.228, 101.193, 21.649]
  MoveL 212 to (-400.87, -591.56, 1195.72) mm, rotated rx 133.78 ry 32.23 rz -154.85 deg; joints [-44.658, 96.97, -166.2, 155.938, -56.848, 47.556, 1383.279, 91.662, 61.038]
  MoveL 213 to (-447.44, -590.25, 1195.98) mm, rotated rx 135.87 ry 31.57 rz -153.98 deg; joints [-44.658, 96.707, -165.848, 156.176, -55.081, 46.59, 1333.576, 98.813, 43.206]
  MoveL 214 to (-498.72, -589.2, 1195.72) mm, rotated rx 138.74 ry 30.18 rz -152.35 deg; joints [-44.658, 96.655, -165.778, 155.89, -52.463, 45.673, 1283.852, 108.8, 19.418]
  MoveL 215 to (-560.72, -587.9, 1194.15) mm, rotated rx 138.79 ry 30.27 rz -152.44 deg; joints [-44.658, 96.577, -165.777, 156.086, -52.555, 45.483, 1220.948, 110.795, 20.377]
  MoveL 216 to (-639.47, -586.59, 1191.27) mm, rotated rx 142.52 ry 28.36 rz -150.48 deg; joints [-44.658, 97.182, -165.778, 155.693, -48.537, 44.439, 1141.12, 123.686, 0.003]
  MoveL 217 to (-727.63, -585.28, 1187.35) mm, rotated rx 144.41 ry 28.4 rz -150.44 deg; joints [-44.658, 97.542, -165.778, 157.123, -47.116, 42.604, 1041.244, 132.367, 0]
  MoveL 218 to (-817.62, -583.97, 1182.38) mm, rotated rx 148.91 ry 26.35 rz -148.6 deg; joints [-44.658, 99.834, -165.778, 156.95, -41.027, 41.319, 939.186, 145.924, 0]
  MoveL 219 to (-903.96, -583.19, 1176.36) mm, rotated rx 152.23 ry 24.86 rz -147.42 deg; joints [-44.738, 101.191, -165.778, 157.354, -36.865, 39.797, 845.179, 158.585, 0]
  MoveL 220 to (-980.87, -582.4, 1170.35) mm, rotated rx 154.34 ry 24.33 rz -146.96 deg; joints [-44.991, 101.599, -165.778, 158.922, -34.925, 37.667, 763.465, 166.916, 0]
  MoveL 221 to (-1045.23, -582.4, 1163.81) mm, rotated rx 157.67 ry 23.31 rz -146.16 deg; joints [-45.554, 102.479, -165.778, 161.669, -31.573, 34.101, 693.904, 177.207, 0]
  MoveL 222 to (-1093.1, -582.92, 1158.31) mm, rotated rx 160.05 ry 23.09 rz -145.83 deg; joints [-46.103, 102.703, -165.778, 165.192, -30.035, 30.105, 641.266, 183.81, 0]
  MoveL 223 to (-1127.38, -584.23, 1152.56) mm, rotated rx 159.19 ry 26.94 rz -147.87 deg; joints [-46.079, 100.059, -165.778, 170.003, -36.283, 26.091, 589.59, 183.81, 2.206]
  MoveL 224 to (-1150.66, -587.37, 1144.71) mm, rotated rx 155.94 ry 32.75 rz -152.02 deg; joints [-44.701, 99.059, -165.778, 172.164, -43.641, 25.274, 521.216, 184.543, 49.963]
  MoveL 225 to (-1167.93, -592.34, 1135.03) mm, rotated rx 153.43 ry 35.4 rz -154.59 deg; joints [-44.467, 96.744, -165.778, 173.427, -49.156, 25.326, 497.205, 184.543, 59.438]
  MoveL 226 to (-1183.88, -598.62, 1122.99) mm, rotated rx 151.57 ry 36.93 rz -156.37 deg; joints [-44.467, 94.397, -165.778, 174.26, -53.492, 25.506, 484.107, 184.541, 61.401]
  MoveL 227 to (-1198.01, -605.42, 1109.65) mm, rotated rx 148.78 ry 38.82 rz -158.96 deg; joints [-44.467, 91.959, -165.778, 175.138, -58.582, 26.153, 472.468, 184.54, 70.526]
  MoveL 228 to (-1209.26, -611.7, 1097.36) mm, rotated rx 147 ry 39.68 rz -160.44 deg; joints [-44.467, 90.097, -165.778, 175.416, -61.854, 26.747, 467.28, 184.54, 74.718]
  MoveL 229 to (-1219.72, -617.98, 1084.54) mm, rotated rx 144.88 ry 40.67 rz -162.27 deg; joints [-44.467, 88.389, -165.778, 175.791, -65.216, 27.456, 461.504, 184.539, 83.939]
  MoveL 230 to (-1231.24, -625.31, 1069.36) mm, rotated rx 143.52 ry 41.13 rz -163.31 deg; joints [-44.467, 86.674, -165.778, 175.885, -67.847, 27.962, 458.129, 184.539, 89.097]
  MoveL 231 to (-1243.79, -633.42, 1051.83) mm, rotated rx 141.86 ry 41.19 rz -164.05 deg; joints [-44.792, 85.593, -165.778, 175.682, -69.649, 28.964, 458.127, 174.356, 102.09]
  MoveL 232 to (-1258.18, -643.1, 1031.17) mm, rotated rx 140.7 ry 41.25 rz -164.59 deg; joints [-45.169, 84.091, -165.778, 175.755, -71.675, 29.544, 458.127, 166.68, 112.151]
  MoveL 233 to (-1272.83, -653.3, 1008.67) mm, rotated rx 138.47 ry 42.09 rz -166.6 deg; joints [-45.169, 82.243, -165.778, 176.203, -75.155, 30.26, 450.031, 166.68, 131.186]
  MoveL 234 to (-1285.91, -663.76, 985.65) mm, rotated rx 135.1 ry 43.09 rz -169.56 deg; joints [-45.169, 80.415, -165.778, 176.756, -79.265, 31.488, 442.666, 166.68, 157.811]
  MoveL 235 to (-1296.12, -673.97, 963.41) mm, rotated rx 132.2 ry 43.79 rz -172.12 deg; joints [-45.169, 78.832, -165.778, 177.232, -82.712, 32.573, 438.161, 166.68, 182.703]
  MoveL 236 to (-1301.61, -683.38, 943) mm, rotated rx 127.99 ry 44.17 rz -175.11 deg; joints [-45.438, 78.266, -165.778, 177.474, -85.57, 34.55, 438.159, 155.427, 220.19]
  MoveL 237 to (-1303.18, -692.02, 924.17) mm, rotated rx 122.92 ry 44.25 rz -178.39 deg; joints [-45.438, 79.694, -167.696, 177.195, -88.679, 37.059, 439.218, 142.971, 279.233]
  MoveL 238 to (-1301.87, -700.13, 907.16) mm, rotated rx 119.59 ry 44.04 rz 179.85 deg; joints [-45.679, 80.765, -169.148, 176.921, -90.687, 38.814, 447.599, 129.185, 323.312]
  MoveL 239 to (-1298.21, -707.71, 891.2) mm, rotated rx 116.95 ry 43.84 rz 178.45 deg; joints [-45.793, 81.677, -170.393, 176.678, -92.348, 40.182, 456.242, 118.579, 361.788]
  MoveL 240 to (-1292.98, -715.3, 876.03) mm, rotated rx 115.79 ry 43.72 rz 177.91 deg; joints [-45.906, 82.066, -170.927, 176.571, -93.064, 40.796, 464.8, 108.892, 386.659]
  MoveL 241 to (-1286.7, -722.36, 861.9) mm, rotated rx 114.7 ry 43.24 rz 178.49 deg; joints [-47.024, 82.267, -171.179, 176.426, -93.438, 41.67, 490.95, 85.22, 406.365]
  MoveL 242 to (-1279.63, -729.69, 848.04) mm, rotated rx 114.07 ry 43.06 rz 178.56 deg; joints [-47.421, 82.432, -171.406, 176.355, -93.755, 42.093, 505.529, 72.113, 424.568]
  MoveL 243 to (-1272.05, -736.49, 834.7) mm, rotated rx 114.85 ry 43.1 rz 179 deg; joints [-47.361, 82.006, -171.406, 176.355, -93.755, 41.68, 514.409, 69.006, 429.679]
  Set speed (1000.0 mm/s)
  MoveL 244 to (-1272.05, -736.49, 834.7) mm, rotated rx 114.85 ry 43.1 rz 179 deg; joints [-47.361, 82.006, -171.406, 176.355, -93.755, 41.68, 514.409, 69.006, 429.679]
  MoveL 245 to (-1302.34, -826.72, 865.38) mm, rotated rx 114.85 ry 43.1 rz 179 deg; joints [-47.361, 82.006, -171.406, 176.355, -93.755, 41.68, 484.114, -21.221, 398.996]

--- program DoorFL (robot ABB IRB 1300-10/1.15) ---
  Smooth(1)
  Set speed (1000.0 mm/s)
  Set Ref.: DoorFL
  Set Tool: Generic Paint Sprayer
  Show Generic Paint Sprayer
  MoveJ 1 to (1.34, 204.65, 100.32) mm, rotated rx 0.03 ry -2.77 rz 73.31 deg; joints [66.672, -21.904, 5.671, 135.111, -6.589, -62.842, 2832.974, 3452.351, 869.235]
  MoveL 2 to (1.34, 204.65, 100.32) mm, rotated rx 0.03 ry -2.77 rz 73.31 deg; joints [66.672, -21.904, 5.671, 135.111, -6.589, -62.842, 2832.974, 3452.351, 869.235]
  MoveL 3 to (0, 200, 200.2) mm, rotated rx 0.03 ry -2.77 rz 73.31 deg; joints [66.672, -21.904, 5.671, 135.111, -6.589, -62.842, 2831.961, 3352.41, 872.535]
  MoveL 4 to (0, 200, 200.2) mm, rotated rx 0.03 ry -2.77 rz 73.31 deg; joints [66.672, -21.904, 5.671, 135.111, -6.589, -62.842, 2831.961, 3352.41, 872.535]
  Set speed (20.0 mm/s)
  MoveL 5 to (0, 100, 183.78) mm, rotated rx -80.27 ry -22.7 rz 88.5 deg; joints [66.672, 3.138, 5.671, 25.397, -90.341, 93.659, 2831.961, 3116.026, 609.959]
  MoveL 6 to (0, 0, 148.68) mm, rotated rx -37.2 ry -3.97 rz 93.93 deg; joints [18.254, 14.754, 0, -34.776, -57.174, 152.551, 2457.292, 3204.962, 879.784]
  Set speed (1000.0 mm/s)
  MoveL 7 to (0, 0, 148.68) mm, rotated rx -37.2 ry -3.97 rz 93.93 deg; joints [18.254, 14.754, 0, -34.776, -57.174, 152.551, 2457.292, 3204.962, 879.784]
  MoveL 8 to (59.94, 9.65, 69.22) mm, rotated rx -37.2 ry -3.97 rz 93.93 deg; joints [18.254, 14.754, 0, -34.776, -57.174, 152.551, 2455.593, 3283.611, 818.047]
  Set speed (1000.0 mm/s)
  MoveL 9 to (75.68, 3.8, 93.4) mm, rotated rx -0.52 ry -2.15 rz 93.34 deg; joints [11.045, 14.885, 0.919, -75.579, -52.247, 159.489, 2455.593, 3283.611, 1100]
  MoveL 10 to (75, 0, 193.33) mm, rotated rx -0.52 ry -2.15 rz 93.34 deg; joints [11.045, 14.656, 0.873, -75.785, -52.179, 159.825, 2455.593, 3183.306, 1100]
  MoveL 11 to (75, 0, 193.33) mm, rotated rx -0.52 ry -2.15 rz 93.34 deg; joints [11.045, 14.656, 0.873, -75.785, -52.179, 159.825, 2455.593, 3183.306, 1100]
  Set speed (20.0 mm/s)
  MoveL 12 to (75, 100, 197.08) mm, rotated rx -0.75 ry -2.14 rz 93.33 deg; joints [11.045, 14.629, 0.873, -75.567, -52.252, 159.825, 2356.015, 3184.966, 1091.846]
  Set speed (1000.0 mm/s)

--- program DoorRL (robot ABB IRB 1300-10/1.15) ---
  Smooth(1)
  Set speed (1000.0 mm/s)
  Set Ref.: DoorRL
  Set Tool: Generic Paint Sprayer
  Show Generic Paint Sprayer
  MoveJ 1 to (98.77, -0.89, 136.35) mm, rotated rx -81.03 ry 0.62 rz 89.58 deg; joints [86.452, 17.717, 3.912, 207.638, 95.308, -83.342, 2064.306, 3452.351, 635.676]
  MoveL 2 to (98.77, -0.89, 136.35) mm, rotated rx -81.03 ry 0.62 rz 89.58 deg; joints [86.452, 17.717, 3.912, 207.638, 95.308, -83.342, 2064.306, 3452.351, 635.676]
  MoveL 3 to (0, 0, 151.94) mm, rotated rx -81.03 ry 0.62 rz 89.58 deg; joints [86.773, 22.351, 7.079, 208.306, 102.336, -79.9, 2064.306, 3452.351, 803.193]
  MoveL 4 to (0, 0, 151.94) mm, rotated rx -81.03 ry 0.62 rz 89.58 deg; joints [86.773, 22.351, 7.079, 208.306, 102.336, -79.9, 2064.306, 3452.351, 803.193]
  Set speed (20.0 mm/s)
  MoveL 5 to (0, 100, 145.88) mm, rotated rx -81.66 ry 0.61 rz 89.52 deg; joints [94.292, 22.53, 7.245, 210.621, 106.407, -85.299, 2064.306, 3452.351, 803.193]
  MoveL 6 to (0, 200, 137.65) mm, rotated rx -81.83 ry 0.63 rz 89.38 deg; joints [101.709, 23.296, 6.366, 212.333, 109.834, -91.105, 2064.306, 3452.351, 803.193]
  Set speed (1000.0 mm/s)
  MoveL 7 to (0, 200, 137.65) mm, rotated rx -81.83 ry 0.63 rz 89.38 deg; joints [101.709, 23.296, 6.366, 212.333, 109.834, -91.105, 2064.306, 3452.351, 803.193]
  MoveL 8 to (98.98, 198.77, 123.44) mm, rotated rx -81.83 ry 0.63 rz 89.38 deg; joints [101.825, 26.359, 16.549, 215.901, 120.872, -82.981, 2064.306, 3452.351, 803.193]
